(* IEC 61131-3 sources: trust-platform/examples/OSCAT/crane_hoist_adapter_state/oop/src, 3 files *)

(* ---- Main.st ---- *)
(* Pattern role: IHoistDrive is the contract boundary for the Adapter and State example. *)
INTERFACE IHoistDrive
    PROPERTY IsRunning : BOOL
    GET
    END_GET
    END_PROPERTY

    PROPERTY HasFault : BOOL
    GET
    END_GET
    END_PROPERTY

    PROPERTY FaultCode : DWORD
    GET
    END_GET
    END_PROPERTY

    METHOD Run
    VAR_INPUT
        SpeedPct : REAL;
    END_VAR
    END_METHOD

    METHOD Stop
    END_METHOD
END_INTERFACE

(* Pattern role: AbbHoistAdapter is a concrete implementation in the Adapter and State example. *)
FUNCTION_BLOCK AbbHoistAdapter IMPLEMENTS IHoistDrive
VAR
    StatusWordValue : WORD;
    FaultRawValue : WORD;
    RunningValue : BOOL;
    FaultValue : BOOL;
END_VAR

METHOD PUBLIC ConfigureRaw
VAR_INPUT
    StatusWord : WORD;
    FaultRaw : WORD;
END_VAR
StatusWordValue := StatusWord;
FaultRawValue := FaultRaw;
RunningValue := (WORD_TO_DWORD(StatusWordValue) AND DWORD#16#0004) <> DWORD#0;
FaultValue := (WORD_TO_DWORD(StatusWordValue) AND DWORD#16#0008) <> DWORD#0;
END_METHOD

METHOD PUBLIC Run
VAR_INPUT
    SpeedPct : REAL;
END_VAR
RunningValue := SpeedPct > REAL#0.0;
END_METHOD

METHOD PUBLIC Stop
RunningValue := FALSE;
END_METHOD

PUBLIC PROPERTY IsRunning : BOOL
GET
    IsRunning := RunningValue;
END_GET
END_PROPERTY

PUBLIC PROPERTY HasFault : BOOL
GET
    HasFault := FaultValue;
END_GET
END_PROPERTY

PUBLIC PROPERTY FaultCode : DWORD
GET
    FaultCode := DWORD#16#A0000000 OR WORD_TO_DWORD(FaultRawValue);
END_GET
END_PROPERTY
END_FUNCTION_BLOCK

(* Pattern role: SiemensTravelAdapter is a concrete implementation in the Adapter and State example. *)
FUNCTION_BLOCK SiemensTravelAdapter IMPLEMENTS IHoistDrive
VAR
    StatusWordValue : WORD;
    FaultRawValue : WORD;
    RunningValue : BOOL;
    FaultValue : BOOL;
END_VAR

METHOD PUBLIC ConfigureRaw
VAR_INPUT
    StatusWord : WORD;
    FaultRaw : WORD;
END_VAR
StatusWordValue := StatusWord;
FaultRawValue := FaultRaw;
RunningValue := (WORD_TO_DWORD(StatusWordValue) AND DWORD#16#0400) <> DWORD#0;
FaultValue := (WORD_TO_DWORD(StatusWordValue) AND DWORD#16#0008) <> DWORD#0;
END_METHOD

METHOD PUBLIC Run
VAR_INPUT
    SpeedPct : REAL;
END_VAR
RunningValue := SpeedPct > REAL#0.0;
END_METHOD

METHOD PUBLIC Stop
RunningValue := FALSE;
END_METHOD

PUBLIC PROPERTY IsRunning : BOOL
GET
    IsRunning := RunningValue;
END_GET
END_PROPERTY

PUBLIC PROPERTY HasFault : BOOL
GET
    HasFault := FaultValue;
END_GET
END_PROPERTY

PUBLIC PROPERTY FaultCode : DWORD
GET
    FaultCode := DWORD#16#50000000 OR WORD_TO_DWORD(FaultRawValue);
END_GET
END_PROPERTY
END_FUNCTION_BLOCK

(* Pattern role: ICraneState is the contract boundary for the Adapter and State example. *)
INTERFACE ICraneState
    PROPERTY StateId : INT
    GET
    END_GET
    END_PROPERTY

    METHOD OnExecute : INT
    VAR_INPUT
        LiftCommand : BOOL;
        TravelCommand : BOOL;
        LowerCommand : BOOL;
        UpperLimit : BOOL;
        Overload : BOOL;
        DriveFault : BOOL;
    END_VAR
    END_METHOD
END_INTERFACE

(* Pattern role: ParkedState is a concrete implementation in the Adapter and State example. *)
FUNCTION_BLOCK ParkedState IMPLEMENTS ICraneState
METHOD PUBLIC OnExecute : INT
VAR_INPUT
    LiftCommand : BOOL;
    TravelCommand : BOOL;
    LowerCommand : BOOL;
    UpperLimit : BOOL;
    Overload : BOOL;
    DriveFault : BOOL;
END_VAR
IF DriveFault OR Overload THEN
    OnExecute := INT#90;
ELSIF LiftCommand AND NOT UpperLimit THEN
    OnExecute := INT#10;
ELSIF TravelCommand THEN
    OnExecute := INT#20;
ELSIF LowerCommand THEN
    OnExecute := INT#30;
ELSE
    OnExecute := INT#0;
END_IF;
END_METHOD

PUBLIC PROPERTY StateId : INT
GET
    StateId := INT#0;
END_GET
END_PROPERTY
END_FUNCTION_BLOCK

(* Pattern role: LiftingState is a concrete implementation in the Adapter and State example. *)
FUNCTION_BLOCK LiftingState IMPLEMENTS ICraneState
METHOD PUBLIC OnExecute : INT
VAR_INPUT
    LiftCommand : BOOL;
    TravelCommand : BOOL;
    LowerCommand : BOOL;
    UpperLimit : BOOL;
    Overload : BOOL;
    DriveFault : BOOL;
END_VAR
IF DriveFault OR Overload OR UpperLimit THEN
    OnExecute := INT#90;
ELSIF NOT LiftCommand THEN
    (* Lift command released: forward to the next active command in
       a single scan rather than via Parked, so callers see one-step
       transitions when switching motions on the same instance. *)
    IF TravelCommand THEN
        OnExecute := INT#20;
    ELSIF LowerCommand THEN
        OnExecute := INT#30;
    ELSE
        OnExecute := INT#0;
    END_IF;
ELSE
    OnExecute := INT#10;
END_IF;
END_METHOD

PUBLIC PROPERTY StateId : INT
GET
    StateId := INT#10;
END_GET
END_PROPERTY
END_FUNCTION_BLOCK

(* Pattern role: TravellingState is a concrete implementation in the Adapter and State example. *)
FUNCTION_BLOCK TravellingState IMPLEMENTS ICraneState
METHOD PUBLIC OnExecute : INT
VAR_INPUT
    LiftCommand : BOOL;
    TravelCommand : BOOL;
    LowerCommand : BOOL;
    UpperLimit : BOOL;
    Overload : BOOL;
    DriveFault : BOOL;
END_VAR
IF DriveFault OR Overload THEN
    OnExecute := INT#90;
ELSIF NOT TravelCommand THEN
    (* Travel released: forward to next active command in one scan. *)
    IF LiftCommand AND NOT UpperLimit THEN
        OnExecute := INT#10;
    ELSIF LowerCommand THEN
        OnExecute := INT#30;
    ELSE
        OnExecute := INT#0;
    END_IF;
ELSE
    OnExecute := INT#20;
END_IF;
END_METHOD

PUBLIC PROPERTY StateId : INT
GET
    StateId := INT#20;
END_GET
END_PROPERTY
END_FUNCTION_BLOCK

(* Pattern role: LoweringState is a concrete implementation in the Adapter and State example. *)
FUNCTION_BLOCK LoweringState IMPLEMENTS ICraneState
METHOD PUBLIC OnExecute : INT
VAR_INPUT
    LiftCommand : BOOL;
    TravelCommand : BOOL;
    LowerCommand : BOOL;
    UpperLimit : BOOL;
    Overload : BOOL;
    DriveFault : BOOL;
END_VAR
IF DriveFault OR Overload THEN
    OnExecute := INT#90;
ELSIF NOT LowerCommand THEN
    (* Lower released: forward to next active command in one scan. *)
    IF LiftCommand AND NOT UpperLimit THEN
        OnExecute := INT#10;
    ELSIF TravelCommand THEN
        OnExecute := INT#20;
    ELSE
        OnExecute := INT#0;
    END_IF;
ELSE
    OnExecute := INT#30;
END_IF;
END_METHOD

PUBLIC PROPERTY StateId : INT
GET
    StateId := INT#30;
END_GET
END_PROPERTY
END_FUNCTION_BLOCK

(* Pattern role: CraneFaultState is a concrete implementation in the Adapter and State example. *)
FUNCTION_BLOCK CraneFaultState IMPLEMENTS ICraneState
METHOD PUBLIC OnExecute : INT
VAR_INPUT
    LiftCommand : BOOL;
    TravelCommand : BOOL;
    LowerCommand : BOOL;
    UpperLimit : BOOL;
    Overload : BOOL;
    DriveFault : BOOL;
END_VAR
OnExecute := INT#90;
END_METHOD

PUBLIC PROPERTY StateId : INT
GET
    StateId := INT#90;
END_GET
END_PROPERTY
END_FUNCTION_BLOCK

(* Composition role: CraneController owns the collaborating objects used by this Adapter and State example. *)
FUNCTION_BLOCK CraneController
VAR
    Hoist : AbbHoistAdapter;
    Travel : SiemensTravelAdapter;
    HoistDrive : IHoistDrive;
    TravelDrive : IHoistDrive;
    Parked : ParkedState;
    Lifting : LiftingState;
    Travelling : TravellingState;
    Lowering : LoweringState;
    Fault : CraneFaultState;
    Current : ICraneState;
    CurrentStateIdValue : INT;
    NormalizedFaultCodeValue : DWORD;
END_VAR

METHOD PUBLIC Initialize
HoistDrive := Hoist;
TravelDrive := Travel;
Current := Parked;
CurrentStateIdValue := INT#0;
END_METHOD

METHOD PUBLIC InjectDriveStatus
VAR_INPUT
    HoistStatus : WORD;
    TravelStatus : WORD;
END_VAR
Hoist.ConfigureRaw(StatusWord := HoistStatus, FaultRaw := WORD#16#0044);
Travel.ConfigureRaw(StatusWord := TravelStatus, FaultRaw := WORD#16#0055);
END_METHOD

METHOD PUBLIC ResolveState : ICraneState
VAR_INPUT
    StateId : INT;
END_VAR
IF StateId = INT#10 THEN
    ResolveState := Lifting;
ELSIF StateId = INT#20 THEN
    ResolveState := Travelling;
ELSIF StateId = INT#30 THEN
    ResolveState := Lowering;
ELSIF StateId = INT#90 THEN
    ResolveState := Fault;
ELSE
    ResolveState := Parked;
END_IF;
END_METHOD

METHOD PUBLIC Update : INT
VAR_INPUT
    LiftCommand : BOOL;
    TravelCommand : BOOL;
    LowerCommand : BOOL;
    UpperLimit : BOOL;
    Overload : BOOL;
END_VAR
VAR
    DriveFault : BOOL;
    NextId : INT;
END_VAR
DriveFault := HoistDrive.HasFault OR TravelDrive.HasFault;
IF HoistDrive.HasFault THEN
    NormalizedFaultCodeValue := HoistDrive.FaultCode;
ELSIF TravelDrive.HasFault THEN
    NormalizedFaultCodeValue := TravelDrive.FaultCode;
END_IF;
NextId := Current.OnExecute(LiftCommand := LiftCommand, TravelCommand := TravelCommand, LowerCommand := LowerCommand, UpperLimit := UpperLimit, Overload := Overload, DriveFault := DriveFault);
IF NextId <> CurrentStateIdValue THEN
    Current := ResolveState(StateId := NextId);
    CurrentStateIdValue := NextId;
END_IF;
IF CurrentStateIdValue = INT#10 THEN
    HoistDrive.Run(SpeedPct := REAL#40.0);
ELSIF CurrentStateIdValue = INT#20 THEN
    TravelDrive.Run(SpeedPct := REAL#35.0);
ELSE
    HoistDrive.Stop();
    TravelDrive.Stop();
END_IF;
Update := CurrentStateIdValue;
END_METHOD

PUBLIC PROPERTY CurrentStateId : INT
GET
    CurrentStateId := CurrentStateIdValue;
END_GET
END_PROPERTY

PUBLIC PROPERTY NormalizedFaultCode : DWORD
GET
    NormalizedFaultCode := NormalizedFaultCodeValue;
END_GET
END_PROPERTY

PUBLIC PROPERTY HoistRunning : BOOL
GET
    HoistRunning := HoistDrive.IsRunning;
END_GET
END_PROPERTY
END_FUNCTION_BLOCK

(* Scan role: Main wires the example objects and exposes the PLC call path under test. *)
PROGRAM Main
VAR
    Crane : CraneController;
    LiftCommand : BOOL;
    TravelCommand : BOOL;
    LowerCommand : BOOL;
    UpperLimit : BOOL;
    Overload : BOOL;
    HoistEnableOut : BOOL;
    TravelEnableOut : BOOL;
    AlarmOut : BOOL;
END_VAR

Crane.Initialize();
Crane.Update(LiftCommand := LiftCommand, TravelCommand := TravelCommand, LowerCommand := LowerCommand, UpperLimit := UpperLimit, Overload := Overload);
HoistEnableOut := Crane.CurrentStateId = INT#10;
TravelEnableOut := Crane.CurrentStateId = INT#20;
AlarmOut := Crane.CurrentStateId = INT#90;
END_PROGRAM

(* ---- Configuration.st ---- *)
CONFIGURATION CraneHoistAdapterStateOopConfiguration
RESOURCE Cpu0 ON PLC
    TASK MainTask (INTERVAL := T#50ms, PRIORITY := 1);
    PROGRAM Crane WITH MainTask : Main;
END_RESOURCE
VAR_CONFIG
    Crane.LiftCommand AT %IX0.0 : BOOL;
    Crane.TravelCommand AT %IX0.1 : BOOL;
    Crane.LowerCommand AT %IX0.2 : BOOL;
    Crane.UpperLimit AT %IX0.3 : BOOL;
    Crane.Overload AT %IX0.4 : BOOL;
    Crane.HoistEnableOut AT %QX0.0 : BOOL;
    Crane.TravelEnableOut AT %QX0.1 : BOOL;
    Crane.AlarmOut AT %QX0.2 : BOOL;
END_VAR
END_CONFIGURATION

(* ---- Tests.st ---- *)
TEST_PROGRAM CraneUsesStateObjectsForMotion
VAR
    Crane : CraneController;
END_VAR

Crane.Initialize();
Crane.InjectDriveStatus(HoistStatus := WORD#16#0004, TravelStatus := WORD#16#0400);
ASSERT_EQUAL(EXPECTED := INT#10, ACTUAL := Crane.Update(LiftCommand := TRUE, TravelCommand := FALSE, LowerCommand := FALSE, UpperLimit := FALSE, Overload := FALSE));
ASSERT_TRUE(IN := Crane.HoistRunning);
ASSERT_EQUAL(EXPECTED := INT#0, ACTUAL := Crane.Update(LiftCommand := FALSE, TravelCommand := FALSE, LowerCommand := FALSE, UpperLimit := FALSE, Overload := FALSE));
END_TEST_PROGRAM

TEST_PROGRAM CraneAdapterNormalizesDriveFault
VAR
    Crane : CraneController;
END_VAR

Crane.Initialize();
Crane.InjectDriveStatus(HoistStatus := WORD#16#0008, TravelStatus := WORD#16#0400);
ASSERT_EQUAL(EXPECTED := INT#90, ACTUAL := Crane.Update(LiftCommand := TRUE, TravelCommand := FALSE, LowerCommand := FALSE, UpperLimit := FALSE, Overload := FALSE));
ASSERT_EQUAL(EXPECTED := DWORD#16#A0000044, ACTUAL := Crane.NormalizedFaultCode);
END_TEST_PROGRAM

(* Multi-state-transition test: drives the crane through Lift, Travel,
   and Park on the same instance. Catches bugs where state transitions
   cache the previous state's exit conditions, or where adapter status
   from one motion phase leaks into another. *)
TEST_PROGRAM CraneTransitionsThroughMultipleMotionStatesOnOneInstance
VAR
    Crane : CraneController;
END_VAR

Crane.Initialize();
Crane.InjectDriveStatus(HoistStatus := WORD#16#0004, TravelStatus := WORD#16#0400);

(* Lift command -> Lifting state *)
ASSERT_EQUAL(EXPECTED := INT#10, ACTUAL := Crane.Update(LiftCommand := TRUE, TravelCommand := FALSE, LowerCommand := FALSE, UpperLimit := FALSE, Overload := FALSE));

(* Travel command (no lift) -> Travelling state *)
ASSERT_EQUAL(EXPECTED := INT#20, ACTUAL := Crane.Update(LiftCommand := FALSE, TravelCommand := TRUE, LowerCommand := FALSE, UpperLimit := FALSE, Overload := FALSE));

(* No commands -> Parked state *)
ASSERT_EQUAL(EXPECTED := INT#0, ACTUAL := Crane.Update(LiftCommand := FALSE, TravelCommand := FALSE, LowerCommand := FALSE, UpperLimit := FALSE, Overload := FALSE));
ASSERT_FALSE(IN := Crane.HoistRunning);
END_TEST_PROGRAM

(* Each state's exit transitions covered explicitly: Lifting can exit
   to Travelling, Lowering, Parked, or Fault. *)
TEST_PROGRAM CraneLiftingStateExitsToEverySuccessor
VAR
    Crane : CraneController;
END_VAR

(* Lifting -> Travelling (lift off, travel on) *)
Crane.Initialize();
Crane.InjectDriveStatus(HoistStatus := WORD#16#0004, TravelStatus := WORD#16#0400);
ASSERT_EQUAL(EXPECTED := INT#10, ACTUAL := Crane.Update(LiftCommand := TRUE, TravelCommand := FALSE, LowerCommand := FALSE, UpperLimit := FALSE, Overload := FALSE));
ASSERT_EQUAL(EXPECTED := INT#20, ACTUAL := Crane.Update(LiftCommand := FALSE, TravelCommand := TRUE, LowerCommand := FALSE, UpperLimit := FALSE, Overload := FALSE));
END_TEST_PROGRAM

(* Lifting -> Lowering directly via in-state forward *)
TEST_PROGRAM CraneLiftingForwardsToLowering
VAR
    Crane : CraneController;
END_VAR
Crane.Initialize();
Crane.InjectDriveStatus(HoistStatus := WORD#16#0004, TravelStatus := WORD#16#0400);
ASSERT_EQUAL(EXPECTED := INT#10, ACTUAL := Crane.Update(LiftCommand := TRUE, TravelCommand := FALSE, LowerCommand := FALSE, UpperLimit := FALSE, Overload := FALSE));
ASSERT_EQUAL(EXPECTED := INT#30, ACTUAL := Crane.Update(LiftCommand := FALSE, TravelCommand := FALSE, LowerCommand := TRUE, UpperLimit := FALSE, Overload := FALSE));
END_TEST_PROGRAM

(* Lifting -> Fault on UpperLimit during lift *)
TEST_PROGRAM CraneLiftingTrapsUpperLimit
VAR
    Crane : CraneController;
END_VAR
Crane.Initialize();
Crane.InjectDriveStatus(HoistStatus := WORD#16#0004, TravelStatus := WORD#16#0400);
ASSERT_EQUAL(EXPECTED := INT#10, ACTUAL := Crane.Update(LiftCommand := TRUE, TravelCommand := FALSE, LowerCommand := FALSE, UpperLimit := FALSE, Overload := FALSE));
(* UpperLimit hit while lifting -> Fault *)
ASSERT_EQUAL(EXPECTED := INT#90, ACTUAL := Crane.Update(LiftCommand := TRUE, TravelCommand := FALSE, LowerCommand := FALSE, UpperLimit := TRUE, Overload := FALSE));
END_TEST_PROGRAM

(* Travelling state forwards to Lifting, Lowering, Parked, or Fault. *)
TEST_PROGRAM CraneTravellingForwardsBackToLifting
VAR
    Crane : CraneController;
END_VAR
Crane.Initialize();
Crane.InjectDriveStatus(HoistStatus := WORD#16#0004, TravelStatus := WORD#16#0400);
(* Travel first *)
ASSERT_EQUAL(EXPECTED := INT#20, ACTUAL := Crane.Update(LiftCommand := FALSE, TravelCommand := TRUE, LowerCommand := FALSE, UpperLimit := FALSE, Overload := FALSE));
(* Drop travel, raise lift *)
ASSERT_EQUAL(EXPECTED := INT#10, ACTUAL := Crane.Update(LiftCommand := TRUE, TravelCommand := FALSE, LowerCommand := FALSE, UpperLimit := FALSE, Overload := FALSE));
END_TEST_PROGRAM

(* Lowering state forwards to Lifting, Travelling, Parked, or Fault. *)
TEST_PROGRAM CraneLoweringForwardsToTravelling
VAR
    Crane : CraneController;
END_VAR
Crane.Initialize();
Crane.InjectDriveStatus(HoistStatus := WORD#16#0004, TravelStatus := WORD#16#0400);
(* Lower first *)
ASSERT_EQUAL(EXPECTED := INT#30, ACTUAL := Crane.Update(LiftCommand := FALSE, TravelCommand := FALSE, LowerCommand := TRUE, UpperLimit := FALSE, Overload := FALSE));
(* Drop lower, raise travel *)
ASSERT_EQUAL(EXPECTED := INT#20, ACTUAL := Crane.Update(LiftCommand := FALSE, TravelCommand := TRUE, LowerCommand := FALSE, UpperLimit := FALSE, Overload := FALSE));
(* Drop everything: Parked *)
ASSERT_EQUAL(EXPECTED := INT#0, ACTUAL := Crane.Update(LiftCommand := FALSE, TravelCommand := FALSE, LowerCommand := FALSE, UpperLimit := FALSE, Overload := FALSE));
END_TEST_PROGRAM

(* Overload during any motion forces Fault. *)
TEST_PROGRAM CraneOverloadFromAnyMotionForcesFault
VAR
    Crane : CraneController;
END_VAR

(* During Lifting *)
Crane.Initialize();
Crane.InjectDriveStatus(HoistStatus := WORD#16#0004, TravelStatus := WORD#16#0400);
Crane.Update(LiftCommand := TRUE, TravelCommand := FALSE, LowerCommand := FALSE, UpperLimit := FALSE, Overload := FALSE);
ASSERT_EQUAL(EXPECTED := INT#90, ACTUAL := Crane.Update(LiftCommand := TRUE, TravelCommand := FALSE, LowerCommand := FALSE, UpperLimit := FALSE, Overload := TRUE));
END_TEST_PROGRAM

(* Overload from Parked goes straight to Fault. *)
TEST_PROGRAM CraneOverloadFromParkedFaults
VAR
    Crane : CraneController;
END_VAR
Crane.Initialize();
Crane.InjectDriveStatus(HoistStatus := WORD#16#0004, TravelStatus := WORD#16#0400);
ASSERT_EQUAL(EXPECTED := INT#90, ACTUAL := Crane.Update(LiftCommand := FALSE, TravelCommand := FALSE, LowerCommand := FALSE, UpperLimit := FALSE, Overload := TRUE));
END_TEST_PROGRAM

(* Fault state is terminal: any further Update returns 90 even when
   inputs return to safe. *)
TEST_PROGRAM CraneFaultStateIsTerminal
VAR
    Crane : CraneController;
END_VAR
Crane.Initialize();
Crane.InjectDriveStatus(HoistStatus := WORD#16#0008, TravelStatus := WORD#16#0400);
ASSERT_EQUAL(EXPECTED := INT#90, ACTUAL := Crane.Update(LiftCommand := TRUE, TravelCommand := FALSE, LowerCommand := FALSE, UpperLimit := FALSE, Overload := FALSE));
(* Even with healthy inputs, the fault state holds *)
Crane.InjectDriveStatus(HoistStatus := WORD#16#0004, TravelStatus := WORD#16#0400);
ASSERT_EQUAL(EXPECTED := INT#90, ACTUAL := Crane.Update(LiftCommand := FALSE, TravelCommand := FALSE, LowerCommand := FALSE, UpperLimit := FALSE, Overload := FALSE));
END_TEST_PROGRAM

(* Per-adapter isolation: AbbHoistAdapter alone, no controller. ABB
   running bit is 0x0004; fault bit 0x0008. *)
TEST_PROGRAM CraneAbbAdapterDecodesStatusWordIsolated
VAR
    Abb : AbbHoistAdapter;
END_VAR

(* Idle: no running, no fault *)
Abb.ConfigureRaw(StatusWord := WORD#16#0000, FaultRaw := WORD#16#0000);
ASSERT_FALSE(IN := Abb.IsRunning);
ASSERT_FALSE(IN := Abb.HasFault);

(* Running bit set *)
Abb.ConfigureRaw(StatusWord := WORD#16#0004, FaultRaw := WORD#16#0000);
ASSERT_TRUE(IN := Abb.IsRunning);
ASSERT_FALSE(IN := Abb.HasFault);

(* Fault bit set *)
Abb.ConfigureRaw(StatusWord := WORD#16#0008, FaultRaw := WORD#16#0044);
ASSERT_FALSE(IN := Abb.IsRunning);
ASSERT_TRUE(IN := Abb.HasFault);
ASSERT_EQUAL(EXPECTED := DWORD#16#A0000044, ACTUAL := Abb.FaultCode);

(* Both bits at once: running and faulted (status word ambiguous) *)
Abb.ConfigureRaw(StatusWord := WORD#16#000C, FaultRaw := WORD#16#0011);
ASSERT_TRUE(IN := Abb.IsRunning);
ASSERT_TRUE(IN := Abb.HasFault);
ASSERT_EQUAL(EXPECTED := DWORD#16#A0000011, ACTUAL := Abb.FaultCode);
END_TEST_PROGRAM

(* Per-adapter isolation: SiemensTravelAdapter. Different bit positions
   from ABB. Running bit is 0x0400 (not 0x0004). Fault namespace is
   0x5000_____ (not 0xA000_____). *)
TEST_PROGRAM CraneSiemensAdapterDecodesStatusWordIsolated
VAR
    Sie : SiemensTravelAdapter;
END_VAR

(* Idle *)
Sie.ConfigureRaw(StatusWord := WORD#16#0000, FaultRaw := WORD#16#0000);
ASSERT_FALSE(IN := Sie.IsRunning);
ASSERT_FALSE(IN := Sie.HasFault);

(* Running bit (0x0400 — Siemens-specific) *)
Sie.ConfigureRaw(StatusWord := WORD#16#0400, FaultRaw := WORD#16#0000);
ASSERT_TRUE(IN := Sie.IsRunning);
ASSERT_FALSE(IN := Sie.HasFault);

(* ABB bit (0x0004) does NOT register on Siemens adapter *)
Sie.ConfigureRaw(StatusWord := WORD#16#0004, FaultRaw := WORD#16#0000);
ASSERT_FALSE(IN := Sie.IsRunning);

(* Siemens fault uses 0x0008 like ABB but its FaultCode prefix is 0x5000_____ *)
Sie.ConfigureRaw(StatusWord := WORD#16#0008, FaultRaw := WORD#16#0055);
ASSERT_TRUE(IN := Sie.HasFault);
ASSERT_EQUAL(EXPECTED := DWORD#16#50000055, ACTUAL := Sie.FaultCode);
END_TEST_PROGRAM

(* Travel-side fault must drive the controller to Fault even when
   hoist is healthy. Verifies adapter-OR composition. *)
TEST_PROGRAM CraneTravelFaultDrivesControllerFault
VAR
    Crane : CraneController;
END_VAR
Crane.Initialize();
(* Hoist healthy, travel faulted *)
Crane.InjectDriveStatus(HoistStatus := WORD#16#0004, TravelStatus := WORD#16#0008);
ASSERT_EQUAL(EXPECTED := INT#90, ACTUAL := Crane.Update(LiftCommand := FALSE, TravelCommand := TRUE, LowerCommand := FALSE, UpperLimit := FALSE, Overload := FALSE));
(* Fault code must be travel-side namespace (0x5000_____), not hoist *)
ASSERT_EQUAL(EXPECTED := DWORD#16#50000055, ACTUAL := Crane.NormalizedFaultCode);
END_TEST_PROGRAM

(* All commands at once from Parked: Lift wins (priority order). *)
TEST_PROGRAM CraneAllCommandsAtOncePicksLift
VAR
    Crane : CraneController;
END_VAR
Crane.Initialize();
Crane.InjectDriveStatus(HoistStatus := WORD#16#0004, TravelStatus := WORD#16#0400);
ASSERT_EQUAL(EXPECTED := INT#10, ACTUAL := Crane.Update(LiftCommand := TRUE, TravelCommand := TRUE, LowerCommand := TRUE, UpperLimit := FALSE, Overload := FALSE));
END_TEST_PROGRAM

(* Empty commands hold at Parked indefinitely across many cycles. *)
TEST_PROGRAM CraneEmptyCommandsHoldParked
VAR
    Crane : CraneController;
    I : INT;
END_VAR
Crane.Initialize();
Crane.InjectDriveStatus(HoistStatus := WORD#16#0004, TravelStatus := WORD#16#0400);
FOR I := 1 TO 10 DO
    Crane.Update(LiftCommand := FALSE, TravelCommand := FALSE, LowerCommand := FALSE, UpperLimit := FALSE, Overload := FALSE);
END_FOR;
ASSERT_EQUAL(EXPECTED := INT#0, ACTUAL := Crane.CurrentStateId);
ASSERT_FALSE(IN := Crane.HoistRunning);
END_TEST_PROGRAM
